// TIA Portal V20 export
// export: Created 2026-10-12T05:06:05.1248225Z, ExportSetting WithDefaults, DisplayName Totally Integrated Automation Portal, DisplayVersion V20, DisplayName TIA Portal Openness, DisplayVersion V20, DisplayName TIA Portal Teamcenter Gateway, DisplayVersion V20, DisplayName TIA Portal Version Control Interface, DisplayVersion V20, DisplayName SINAMICS Startdrive Advanced, DisplayVersion V20 SP1 Update 2, DisplayName SINAMICS Startdrive G110M, G120, G120C, G120D, G120P, G115D, DisplayVersion V20 SP1 Update 2, DisplayName SINAMICS Startdrive G130, G150, S120, S150, SINAMICS MV, G220, S200, S210, DisplayVersion V20 SP1 Update 2, DisplayName STEP 7 Professional, DisplayVersion V20, DisplayName STEP 7 Safety, DisplayVersion V20, DisplayName WinCC Basic/Comfort/Advanced, DisplayVersion V20, DisplayName WinCC Professional, DisplayVersion V20, DisplayName WinCC Unified, DisplayVersion V20
FUNCTION "FRK_SetResult" : Void   // FC117, SCL
{ S7_Optimized_Access := 'TRUE' }
VERSION : 0.1
// stored: AutoNumber true, IsIECCheckEnabled false, SetENOAutomatically false, UDAEnableTagReadback false
   VAR_INPUT
      Request : "ST_HmiRequest";
      Response : "ST_HmiResponse";
      Scope : String;
      RootIndex : Int;
   END_VAR
   VAR_IN_OUT
      Persist : "ST_ConfigPersistStatus";
      AlarmLog : "FRK_AlarmLog";
   END_VAR
   VAR_TEMP
      Diag : "ST_Diagnostic";
      Slot : Int;
      Ok : Bool;
   END_VAR
BEGIN

   IF #Request.Kind <> 29 THEN
       RETURN;
   END_IF;
   IF NOT #Response.Accepted THEN
       #Persist.LastRejectScope := "FRK_SetRuntime".Work[#RootIndex].RejectScope;
       #Persist.LastRejectKey := "FRK_SetRuntime".Work[#RootIndex].RejectKey;
   END_IF;
   #Diag := "FRK_UnitScratch".EmptyDiagnostic;
   #Diag.SourcePath := STRING_TO_WSTRING(#Scope);
   IF #Response.Accepted THEN
       #Diag.ReasonCode := 2043;
       #Diag.Description := WSTRING#'std.event.configSetApplied';
   ELSE
       #Diag.ReasonCode := 2042;
       #Diag.Description := WSTRING#'std.error.configSetRejected';
       #Diag.SourcePath := STRING_TO_WSTRING(#Persist.LastRejectScope);
   END_IF;
   #Slot := "FRK_AlarmRaise"(AlarmLog := #AlarmLog, Diag := #Diag, ResetClass := 0);
   IF #Slot > 0 THEN
       #Ok := "FRK_AlarmGone"(AlarmLog := #AlarmLog, Slot := #Slot);
   END_IF;
END_FUNCTION
